ABB RAPID module: TCP_ProtJSD.mod

MODULE TCP_ProtJSD
	! Points are read in order of declaration.
  ! Please do not change the order of points!

  LOCAL PERS robtarget pTCP_Point1:=[[365.1418,0.135368,667.08],[0.580704092979431,0.0454636663198471,0.812194585800171,0.0324912779033184],[0,-1,0,0],[9E+09,9E+09,9E+09,9E+09,9E+09,9E+09]];
	LOCAL PERS robtarget pTCP_Point2:=[[331.0422,37.52399,622.4653],[0.636924266815186,-0.192049846053123,0.739533483982086,-0.102637745440006],[0,-1,-1,0],[9E+09,9E+09,9E+09,9E+09,9E+09,9E+09]];
	LOCAL PERS robtarget pTCP_Point3:=[[351.9474,-62.10214,635.1849],[0.581058382987976,0.191919669508934,0.771535396575928,0.173985943198204],[-1,0,-1,0],[9E+09,9E+09,9E+09,9E+09,9E+09,9E+09]];
	LOCAL PERS robtarget pTCP_Point4:=[[409.1765,-45.67894,696.2203],[0.511161506175995,-0.16655920445919,0.840345561504364,0.0692193657159805],[-1,0,-1,0],[9E+09,9E+09,9E+09,9E+09,9E+09,9E+09]];

ENDMODULE
